Fanuc KAREL source: kt00514.KL

-- PROVISIONAL review KL for V770-1; original PC SHA256 de3aa1178563fff54d2e9998ab94bdaec641dbfd3a5921de248f58a382eaaecb
-- Incomplete behavior may be omitted. Consult companion uncertainty JSON. Do not deploy.
PROGRAM KT00514
%NOLOCKGROUP
-- UNRESOLVED_DECL P1 type=000106
-- UNRESOLVED_DECL P2 type=000101
-- UNRESOLVED_DECL OUT type=000101
BEGIN
  -- UNRESOLVED_PC offsets 5-20; opcodes 2E,22,32,35
  -- UNRESOLVED_PC offsets 25-54; opcodes 49,7E,49,60,4A
  -- UNRESOLVED_PC offsets 59-63; opcodes 7F
END KT00514
